FUNCTION_BLOCK PUMP_DUTY_SELECT (* Migrated from IEC 61131-3 ST *)
  (* Standard: 61499-2 *)
  (* Version 1.0, 2026-11-06, st2fb *)
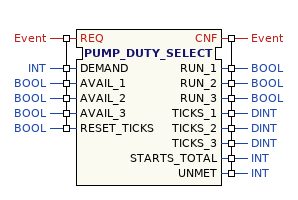
  EVENT_INPUT
    REQ WITH DEMAND, AVAIL_1, AVAIL_2, AVAIL_3, RESET_TICKS;
  END_EVENT
  EVENT_OUTPUT
    CNF WITH RUN_1, RUN_2, RUN_3, TICKS_1, TICKS_2, TICKS_3, STARTS_TOTAL, UNMET;
  END_EVENT
  VAR_INPUT
    DEMAND : INT;
    AVAIL_1 : BOOL;
    AVAIL_2 : BOOL;
    AVAIL_3 : BOOL;
    RESET_TICKS : BOOL;
  END_VAR
  VAR_OUTPUT
    RUN_1 : BOOL;
    RUN_2 : BOOL;
    RUN_3 : BOOL;
    TICKS_1 : DINT;
    TICKS_2 : DINT;
    TICKS_3 : DINT;
    STARTS_TOTAL : INT;
    UNMET : INT;
  END_VAR
  VAR
    PUMP_COUNT : INT := 3;
    WEAR_PER_START : DINT := 5;
    AV1 : BOOL := FALSE;
    AV2 : BOOL := FALSE;
    AV3 : BOOL := FALSE;
    RN1 : BOOL := FALSE;
    RN2 : BOOL := FALSE;
    RN3 : BOOL := FALSE;
    RT1 : DINT := 0;
    RT2 : DINT := 0;
    RT3 : DINT := 0;
    ST1 : INT := 0;
    ST2 : INT := 0;
    ST3 : INT := 0;
    WR1 : BOOL := FALSE;
    WR2 : BOOL := FALSE;
    WR3 : BOOL := FALSE;
    PREV_DEMAND : INT := 0;
    N : INT := 0;
    P : INT := 0;
    BEST : INT := 0;
    BEST_SCORE : DINT := 0;
    SCORE : DINT := 0;
    CHANGED : BOOL := FALSE;
    TMP_B : BOOL := FALSE;
    TMP_A : BOOL := FALSE;
    TMP_D : DINT := 0;
    TMP_I : INT := 0;
    DONE_F : BOOL := FALSE;
  END_VAR
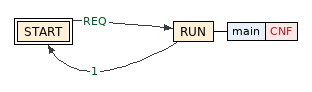
  EC_STATES
    START;
    RUN : main -> CNF;
  END_STATES
  EC_TRANSITIONS
    START TO RUN := REQ;
    RUN TO START := 1;
  END_TRANSITIONS
  ALGORITHM main IN ST:
AV1 := AVAIL_1;
AV2 := AVAIL_2;
AV3 := AVAIL_3;

CHANGED := DEMAND <> PREV_DEMAND;
DONE_F := FALSE;
FOR P := 1 TO 3 DO
  IF NOT DONE_F THEN
    TMP_B := FALSE;
    TMP_A := FALSE;
    IF P = 1 THEN
      TMP_B := RN1;
      TMP_A := AV1;
    ELSIF P = 2 THEN
      TMP_B := RN2;
      TMP_A := AV2;
    ELSE
      TMP_B := RN3;
      TMP_A := AV3;
    END_IF;
    IF TMP_B AND NOT TMP_A THEN
      CHANGED := TRUE;
      DONE_F := TRUE;
    END_IF;
  END_IF;
END_FOR;
PREV_DEMAND := DEMAND;

IF CHANGED THEN
  WR1 := RN1;
  WR2 := RN2;
  WR3 := RN3;
  RN1 := FALSE;
  RN2 := FALSE;
  RN3 := FALSE;
  UNMET := 0;
  DONE_F := FALSE;
  FOR N := 1 TO DEMAND DO
    IF NOT DONE_F THEN
      BEST := 0;
      BEST_SCORE := 2147483647;
      FOR P := 1 TO 3 DO
        TMP_B := FALSE;
        TMP_D := 0;
        IF P = 1 THEN
          TMP_B := AV1 AND NOT RN1;
          TMP_D := RT1 + WEAR_PER_START * INT_TO_DINT(ST1);
        ELSIF P = 2 THEN
          TMP_B := AV2 AND NOT RN2;
          TMP_D := RT2 + WEAR_PER_START * INT_TO_DINT(ST2);
        ELSE
          TMP_B := AV3 AND NOT RN3;
          TMP_D := RT3 + WEAR_PER_START * INT_TO_DINT(ST3);
        END_IF;
        IF TMP_B THEN
          SCORE := TMP_D;
          IF SCORE < BEST_SCORE THEN
            BEST := P;
            BEST_SCORE := SCORE;
          END_IF;
        END_IF;
      END_FOR;
      IF BEST = 0 THEN
        UNMET := DEMAND - N + 1;
        DONE_F := TRUE;
      ELSE
        TMP_B := FALSE;
        IF BEST = 1 THEN
          RN1 := TRUE;
          TMP_B := NOT WR1;
          IF TMP_B THEN
            ST1 := ST1 + 1;
          END_IF;
        ELSIF BEST = 2 THEN
          RN2 := TRUE;
          TMP_B := NOT WR2;
          IF TMP_B THEN
            ST2 := ST2 + 1;
          END_IF;
        ELSE
          RN3 := TRUE;
          TMP_B := NOT WR3;
          IF TMP_B THEN
            ST3 := ST3 + 1;
          END_IF;
        END_IF;
        IF TMP_B THEN
          STARTS_TOTAL := STARTS_TOTAL + 1;
        END_IF;
      END_IF;
    END_IF;
  END_FOR;
END_IF;

IF RESET_TICKS THEN
  RT1 := 0;
  RT2 := 0;
  RT3 := 0;
ELSE
  IF RN1 THEN
    RT1 := RT1 + 1;
  END_IF;
  IF RN2 THEN
    RT2 := RT2 + 1;
  END_IF;
  IF RN3 THEN
    RT3 := RT3 + 1;
  END_IF;
END_IF;

RUN_1 := RN1;
RUN_2 := RN2;
RUN_3 := RN3;
TICKS_1 := RT1;
TICKS_2 := RT2;
TICKS_3 := RT3;
  END_ALGORITHM
END_FUNCTION_BLOCK
